// TIA Portal V19 export
// export: Created 2026-10-15T09:44:23.06076Z, ExportSetting WithDefaults, DisplayName Totally Integrated Automation Portal, DisplayVersion V19, DisplayName TIA Portal Openness, DisplayVersion V19, DisplayName TIA Portal Version Control Interface, DisplayVersion V19, DisplayName STEP 7 Professional, DisplayVersion V19, DisplayName STEP 7 Safety, DisplayVersion V19, DisplayName WinCC Basic/Comfort/Advanced, DisplayVersion V19, DisplayName WinCC Unified, DisplayVersion V19
FUNCTION "ROLL_TimerOp" : Void   // FC6, SCL
{ S7_Optimized_Access := 'TRUE' }
VERSION : 0.1
// stored: AutoNumber true, IsIECCheckEnabled false, SetENOAutomatically false, UDAEnableTagReadback false
   VAR_INPUT
      Number : Int;
      Operation : Int;   // 0=SE on-delay; 1=SA off-delay; 2=R reset
      Signal : Bool;
      Preset : Word;
   END_VAR
   VAR_TEMP
      base : Int;
      count : Int;
      trigger : Bool;
   END_VAR
BEGIN

   IF (#Number < 0) OR (#Number > 127) THEN
       "ROLL_IO".ConversionFault := TRUE;
       RETURN;
   END_IF;
   IF #Operation = 2 THEN
       IF #Signal THEN
           "ROLL_State".S5Timers[#Number].RemainingMs := 0.0;
           "ROLL_State".S5Timers[#Number].Q := FALSE;
       END_IF;
       RETURN;
   END_IF;
   #trigger := ((#Operation = 0) AND #Signal AND NOT "ROLL_State".S5Timers[#Number].Previous)
   OR ((#Operation = 1) AND NOT #Signal AND "ROLL_State".S5Timers[#Number].Previous);
   IF #trigger THEN
       #count := "ROLL_DecodeBCD"(Value := #Preset);
       #base := WORD_TO_INT(SHR(IN := #Preset AND W#16#F000, N := 12));
       CASE #base OF
           0:
               #base := 10;
           1:
               #base := 100;
           2:
               #base := 1000;
           3:
               #base := 10000;
           ELSE
               #base := 0;
       END_CASE;
       IF (#base = 0) OR (#count < 0) THEN
           "ROLL_IO".ConversionFault := TRUE;
           "ROLL_State".S5Timers[#Number].RemainingMs := 0.0;
           "ROLL_State".S5Timers[#Number].Q := FALSE;
           RETURN;
       END_IF;
       "ROLL_State".S5Timers[#Number].BaseMs := #base;
       "ROLL_State".S5Timers[#Number].RemainingMs := INT_TO_LREAL(#count) * INT_TO_LREAL(#base);
   END_IF;
   "ROLL_State".S5Timers[#Number].Mode := #Operation;
   IF #Operation = 0 THEN
       IF NOT #Signal THEN
           "ROLL_State".S5Timers[#Number].RemainingMs := 0.0;
       END_IF;
       "ROLL_State".S5Timers[#Number].Q := #Signal AND ("ROLL_State".S5Timers[#Number].RemainingMs <= 0.0);
   ELSIF #Operation = 1 THEN
       IF #Signal THEN
           "ROLL_State".S5Timers[#Number].RemainingMs := 0.0;
       END_IF;
       "ROLL_State".S5Timers[#Number].Q := #Signal OR ("ROLL_State".S5Timers[#Number].RemainingMs > 0.0);
   ELSE
       "ROLL_IO".ConversionFault := TRUE;
   END_IF;
   "ROLL_State".S5Timers[#Number].Previous := #Signal;
END_FUNCTION
